(* IEC 61131-3 sources: plc-process-lib/src/POUs/Util/FB_LimitMonitor, 2 files *)

(* ---- FB_LimitMonitor.decl.st ---- *)
// Назначение: одна уставка с гистерезисом, задержками срабатывания и снятия и
//             разрешением. Верхняя: флаг при значении >= уставки, снятие ниже уставки минус
//             гистерезис; нижняя — зеркально. Неконечное значение флаг не меняет. Выключенная
//             уставка или xForceOff снимают флаг сразу, без задержки.
// Автор:      kr0nsch
// Версия:     0.1.0
// Документ:   docs/fb/FB_LimitMonitor.md
FUNCTION_BLOCK FB_LimitMonitor
VAR_INPUT
    rValue_eu  : REAL;             // контролируемое значение
    xHighLimit : BOOL;             // TRUE — верхняя уставка (HH, H), FALSE — нижняя (L, LL)
    xForceOff  : BOOL;             // TRUE — флаг FALSE сразу (отказ сигнала, OOS)
    stCfg      : ST_AiLimitCfg;    // параметры уставки
    itfTime    : I_TimeSource;     // источник времени; 0 — встроенный fbSysTime
END_VAR
VAR_OUTPUT
    xOut : BOOL;                   // после гистерезиса и задержек
    xRaw : BOOL;                   // после гистерезиса, до задержек
END_VAR
VAR
    fbDelay   : FB_Delay;          // задержки срабатывания и снятия флага
    fbSysTime : FB_SystemTime;     // запасной источник времени
END_VAR
VAR_TEMP
    itfTimeAct : I_TimeSource;     // действующий источник этого вызова
    xNewRaw    : BOOL;             // флаг после гистерезиса для конечного значения
END_VAR

(* ---- FB_LimitMonitor.impl.st ---- *)
IF NOT stCfg.xEnable OR xForceOff THEN
    // уставка выключена или принудительный сброс: флаг снимается сразу, отсчёт задержек —
    // заново после включения
    xRaw := FALSE;
    fbDelay.Preset(xValue := FALSE);
    xOut := FALSE;
ELSE
    IF itfTime <> 0 THEN
        itfTimeAct := itfTime;
    ELSE
        itfTimeAct := fbSysTime;
    END_IF

    // гистерезис: в зоне между порогами срабатывания и снятия флаг сохраняется
    IF xHighLimit THEN
        xNewRaw := (rValue_eu >= stCfg.rSetpoint_eu)
                   OR (xRaw AND (rValue_eu >= stCfg.rSetpoint_eu - stCfg.rHyst_eu));
    ELSE
        xNewRaw := (rValue_eu <= stCfg.rSetpoint_eu)
                   OR (xRaw AND (rValue_eu <= stCfg.rSetpoint_eu + stCfg.rHyst_eu));
    END_IF
    // неконечное значение (NaN, ±Inf, мусор) флаг не меняет
    xRaw := SEL(F_IsFinite(rIn := rValue_eu), xRaw, xNewRaw);

    fbDelay(xIn := xRaw, tOnDelay := stCfg.tOnDelay, tOffDelay := stCfg.tOffDelay, itfTime := itfTimeAct);
    xOut := fbDelay.xOut;
END_IF
